FUNCTION_BLOCK "naut_Main"
{ S7_Optimized_Access := 'TRUE' }
VERSION : 0.1
   VAR
      count : INT;
      pulse : R_TRIG;
      dwell : TON_TIME;
      naut_dwell_last : Struct
         Q : Bool;
         ET : Time;
      END_STRUCT;
      batches : IEC_LCOUNTER;
      state : INT := 0;
      avg : REAL;
   END_VAR
   VAR RETAIN
      total : DINT;
   END_VAR
   VAR_TEMP
      i : INT;
      naut_for_v1 : INT;
   END_VAR

BEGIN
	#i := 0;
	"naut_Tags".Heartbeat := LINT_TO_UINT(((UINT_TO_LINT("naut_Tags".Heartbeat) + 1) MOD LINT#65536 + LINT#65536) MOD LINT#65536);
	"naut_Tags".Echo := "naut_Tags".Command;
	#pulse(CLK := "naut_Tags".Start);
	#dwell(IN := "naut_Tags".Running AND NOT "naut_Tags".Fault, PT := T#2s, Q => #naut_dwell_last.Q, ET => #naut_dwell_last.ET);
	#batches.CTU(CU := #pulse.Q, R := "naut_Tags".Reset, PV := 10);
	"naut_Tags".Done := #batches.QU;
	IF #naut_dwell_last.Q THEN
		#count := LINT_TO_INT((((INT_TO_LINT(#count) + 1) + LINT#32768) MOD LINT#65536 + LINT#65536) MOD LINT#65536 - LINT#32768);
		#total := LINT_TO_DINT((((DINT_TO_LINT(#total) + DINT_TO_LINT(INT_TO_DINT(#count))) + LINT#2147483648) MOD LINT#4294967296 + LINT#4294967296) MOD LINT#4294967296 - LINT#2147483648);
	ELSIF "naut_Tags".Fault THEN
		#count := 0;
	ELSE
		#count := MIN(IN1 := #count, IN2 := 100);
	END_IF;
	CASE #state OF
		0:
			IF "naut_Tags".Start THEN
				#state := 1;
			END_IF;
		1, 2:
			#state := LINT_TO_INT((((INT_TO_LINT(#state) + 1) + LINT#32768) MOD LINT#65536 + LINT#65536) MOD LINT#65536 - LINT#32768);
		3..5:
			#state := 0;
		ELSE
			#state := 0;
	END_CASE;
	#avg := 0.0;
	FOR #naut_for_v1 := 1 TO 4 DO
		#i := #naut_for_v1;
		#avg := #avg + INT_TO_REAL(#i) / 4.0;
	END_FOR;
	#i := 5;
	"naut_Tags".Level := LIMIT(MN := 0.0, IN := "naut_Tags".Level * 1.5 - (#avg + 2.0), MX := 100.0);
	"naut_Tags".Running := NOT ("naut_Tags".Fault OR "naut_Tags".Reset) AND "naut_Tags".Start;
END_FUNCTION_BLOCK
